(* IEC 61131-3 sources: codesys-framework/txt/application/WeVe Core (library)/10 Mode/FB_Mode, 11 files *)

(* ---- Active.prop.st ---- *)
PROPERTY Active : BOOL

// --- BEGIN IMPLEMENTATION ---

// ----------- SET -----------
VAR
END_VAR

// -- BEGIN IMPLEMENTATION SET --
_xActive := Active;

// ----------- GET -----------
VAR
END_VAR

// -- BEGIN IMPLEMENTATION GET --
Active := _xActive;

(* ---- FB_Init.method.st ---- *)
//FB_Init is always available implicitly and it is used primarily for initialization.
//The return value is not evaluated. For a specific influence, you can also declare the
//methods explicitly and provide additional code there with the standard initialization
//code. You can evaluate the return value.
METHOD FB_Init: BOOL
VAR_INPUT
    bInitRetains: BOOL := TRUE; // TRUE: the retain variables are initialized (reset warm / reset cold)
    bInCopyCode: BOOL := TRUE;  // TRUE: the instance will be copied to the copy code afterward (online change)

	nMode 					: USINT;
	sName 					: STRING;
	fbEventSrv 				: I_EventService;
	fbSafetySrv				: I_SafetyService;
	fbEvents 				: I_EventGroup;		// de gedeelde FB_ModeEventGroup, mag 0 zijn
END_VAR

// --- BEGIN IMPLEMENTATION ---

// Enkel referenties en waarden bewaren, geen methodes aanroepen
_fbEventSrv 	:= fbEventSrv;
_fbSafetySrv 	:= fbSafetySrv;
_fbEvents 		:= fbEvents;

_nMode := nMode;
_sName := sName;

(* ---- InitRequest.method.st ---- *)
METHOD InitRequest

// --- BEGIN IMPLEMENTATION ---

IF _eState = E_ModeStates.Standby THEN
	_eState := E_ModeStates.Initialize;
END_IF

(* ---- Mode.prop.st ---- *)
PROPERTY Mode : USINT

// --- BEGIN IMPLEMENTATION ---

// ----------- GET -----------
VAR
END_VAR

// -- BEGIN IMPLEMENTATION GET --
Mode := _nMode;

(* ---- Name.prop.st ---- *)
PROPERTY Name : STRING
// --- BEGIN IMPLEMENTATION ---

// ----------- GET -----------
VAR
END_VAR

// -- BEGIN IMPLEMENTATION GET --
Name := _sName;

(* ---- ResetEvents.method.st ---- *)
// Alle events van de machine resetten via de EventService (ook die van deze mode).
// Elk event beslist zelf of het mag (conditie weg).
// TRUE = geen enkel event nog actief.
METHOD ResetEvents : BOOL
VAR_INPUT
END_VAR

// --- BEGIN IMPLEMENTATION ---

IF _fbEventSrv <> 0 THEN
	ResetEvents := _fbEventSrv.Reset();
ELSE
	ResetEvents := TRUE;
END_IF

(* ---- ResetSequenceRequest.method.st ---- *)
// TRUE = aanvraag aanvaard.
METHOD ResetSequenceRequest : BOOL
VAR
	scPayload 	: SC_EventPayload;
END_VAR

// --- BEGIN IMPLEMENTATION ---

IF
	_eState = E_ModeStates.Run OR
	_eState = E_ModeStates.Stop OR
	_eState = E_ModeStates.QuickStop
THEN
	IF _fbEvents <> 0 THEN
		scPayload.asPayload[0] := _sName;
		_fbEvents.Log(iEvent := E_ModeEvents.ResetRequestInvalid, scPayload := scPayload);
	END_IF

	ResetSequenceRequest := FALSE;
	RETURN;
END_IF

_eState := E_ModeStates.Reset;
ResetSequenceRequest := TRUE;

(* ---- SetRequest.method.st ---- *)
// Basis: geen mode-specifieke aanvragen. Een concrete mode overschrijft deze methode.
// TRUE = aanvraag aanvaard.
METHOD SetRequest : BOOL
VAR_INPUT
	iRequest	: UINT;
	pData		: POINTER TO ARRAY [0..255] OF BYTE := 0;
	pSize		: ULINT := 0;
END_VAR
VAR
	scPayload 	: SC_EventPayload;
END_VAR

// --- BEGIN IMPLEMENTATION ---

IF _fbEvents <> 0 THEN
	scPayload.asPayload[0] := _sName;
	_fbEvents.Log(iEvent := E_ModeEvents.UserRequestInvalid, scPayload := scPayload);
END_IF

SetRequest := FALSE;

(* ---- StartRequest.method.st ---- *)
// Basis: start is niet mogelijk. Een concrete mode die starten toelaat, overschrijft deze methode.
// TRUE = aanvraag aanvaard.
METHOD StartRequest : BOOL
VAR
	scPayload 	: SC_EventPayload;
END_VAR

// --- BEGIN IMPLEMENTATION ---

IF _fbEvents <> 0 THEN
	scPayload.asPayload[0] := _sName;
	_fbEvents.Log(iEvent := E_ModeEvents.StartRequestInvalid, scPayload := scPayload);
END_IF

StartRequest := FALSE;

(* ---- State.prop.st ---- *)
PROPERTY State : E_ModeStates

// --- BEGIN IMPLEMENTATION ---

// ----------- GET -----------
VAR
END_VAR

// -- BEGIN IMPLEMENTATION GET --
State := _eState;

// ----------- SET -----------
VAR
END_VAR

// -- BEGIN IMPLEMENTATION SET --
_eState := State;

(* ---- StopRequest.method.st ---- *)
METHOD StopRequest

// --- BEGIN IMPLEMENTATION ---

IF 		_eState = E_ModeStates.Starting
	OR 	_eState = E_ModeStates.Run
	OR 	_eState = E_ModeStates.Safe
THEN
	_eState := E_ModeStates.Stop;
END_IF
